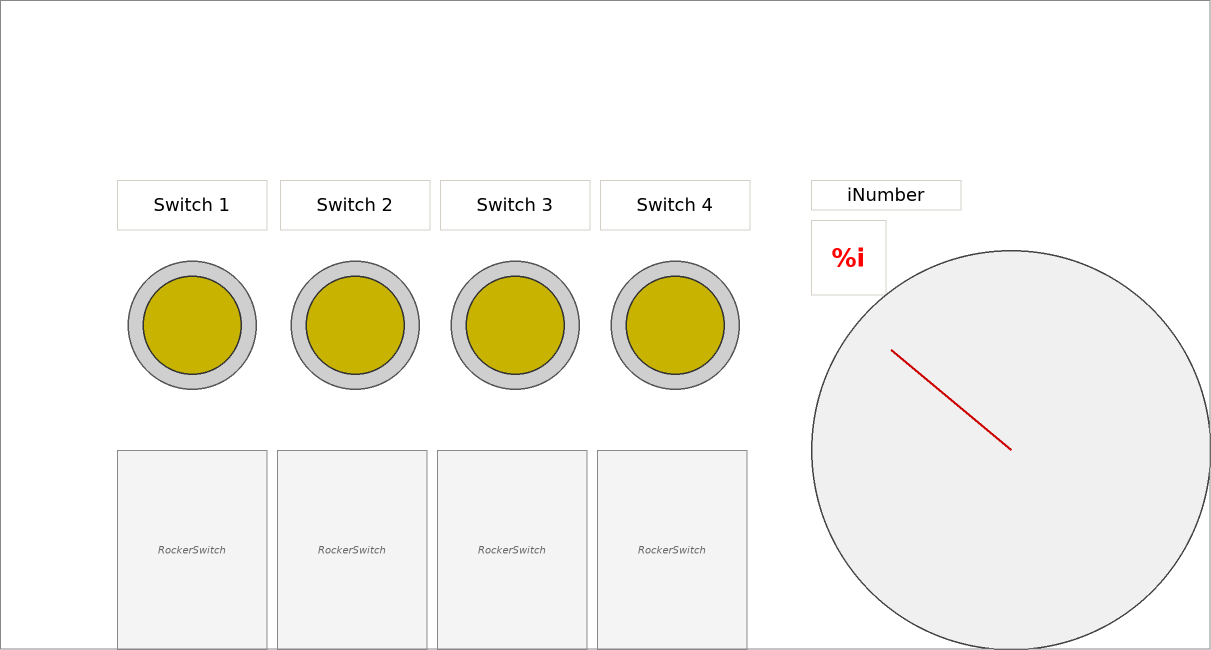
VISUALIZATION Visualization  // 1211x650
    RockerSwitch (117,450 150x200), variable: MAIN.bSwitch1, behaviour: TOGGLE, style: Switch-RockerSwitch-Gray
    RockerSwitch (277,450 150x200), variable: MAIN.bSwitch2, behaviour: TOGGLE, style: Switch-RockerSwitch-Gray
    RockerSwitch (437,450 150x200), variable: MAIN.bSwitch3, behaviour: TOGGLE, style: Switch-RockerSwitch-Gray
    RockerSwitch (597,450 150x200), variable: MAIN.bSwtich4, behaviour: TOGGLE, style: Switch-RockerSwitch-Gray
    Lamp1 (117,250 150x150), variable: MAIN.bLight1, style: Lamp-Lamp1-Yellow
    Lamp1 (440,250 150x150), variable: MAIN.bLight3, style: Lamp-Lamp1-Yellow
    Lamp1 (280,250 150x150), variable: MAIN.bLight2, style: Lamp-Lamp1-Yellow
    Lamp1 (600,250 150x150), variable: MAIN.bLight4, style: Lamp-Lamp1-Yellow
    Textfield (117,180 150x50), "Switch 1"
    Textfield (280,180 150x50), "Switch 2"
    Textfield (440,180 150x50), "Switch 3"
    Textfield (600,180 150x50), "Switch 4"
    Textfield (811,220 75x75), "%i", text variable: MAIN.iNumber
    Textfield (811,180 150x30), "iNumber"
    Meter360 (811,250 400x400), value: MAIN.iNumber, style: Meter-Meter360-Gray, scale format: %.1f, scale 0..32000
END_VISUALIZATION

(* stored: Version 1.1.0.1
   Visu Visualization: Id {032c632f-8b83-4d5f-b4aa-77fdb26114b5} *)
